// TIA Portal project "Text" (V21)

(* hardware
DEVICE "PLC_Text"  S7-1500 station
   slot 0: "Rail_0"  Rack  6ES7 590-1***0-0AA0
   slot 1: "PLC_Text"  CPU 1516-3 PN/DP  6ES7 516-3AN02-0AB0  V2.9
      slot 3: "CPU display_1"  6ES7591-1BA00-0AA0
      slot 32768: "PROFINET interface_1"  X1
         slot 32769: "Port_1"  X1 P1
         slot 32770: "Port_2"  X1 P2
      slot 33024: "PROFINET interface_2"  X2
         slot 33025: "Port_1"  X2 P1
      slot 33280: "DP interface_1"  X3
      slot 34817: "Virtual CP interface port_1"  Virtual CP interface port  Virtual CP interface port
*)

// ===== PLC "PLC_Text"  CPU 1516-3 PN/DP =====

VAR_GLOBAL   // PLC tag table "Beschriftung"
   "Lamp_Überlast" AT %Q0.0 : Bool;   // Überlast der Pumpe – Leuchte
   "Sensor_Niveau" AT %IW2 : Int;   // Capteur de niveau, en ‰
   "Etikett" AT %MW4 : Word;   // ラベル番号 (標識)
END_VAR

TYPE "typeLabel"
   STRUCT
      german : WString[40] := WSTRING#'Füllhöhe überschritten';   // Größe in Millilitern
      french : WString[40] := WSTRING#'Défaut de la vanne';   // Vanne fermée, ça bloque
      japanese : WString[20] := WSTRING#'液面センサー';   // 日本語のコメント
      chinese : WString[20] := WSTRING#'液位传感器';   // 中文注释
      plain : String[20] := 'It$'s 50% full';   // A quote and a percent sign
   END_STRUCT;
END_TYPE

DATA_BLOCK "Labels"   // DB1
TITLE = Beschriftungen für das Bedienfeld
{ S7_Optimized_Access := 'TRUE' }
VERSION : 0.1
   VAR
      current : "typeLabel";   // Die aktuelle Meldung
      list : Array[1..2] of "typeLabel";   // Zur Auswahl
      note : WString[40] := WSTRING#'Notiz: «Anführungszeichen»';   // Guillemets
   END_VAR
BEGIN
   list[1].german := WSTRING#'Ventil öffnet';
   list[2].japanese := WSTRING#'バルブが開く';
END_DATA_BLOCK

FUNCTION_BLOCK "Texts"   // FB1, SCL
TITLE = Überprüfung der Füllhöhe – ½ Liter
{ S7_Optimized_Access := 'TRUE' }
VERSION : 0.1
// Prüft die Füllhöhe. Vérifie le niveau. 液面を確認する。检查液位。
// A second comment line, with symbols: ± ° µ € ✓
   VAR_INPUT
      level : Real;   // Füllhöhe in ml – niveau de remplissage
      limit : Real := 500.0;   // Grenzwert ≥ 0
   END_VAR
   VAR_OUTPUT
      message : WString[60];   // Meldung für das Bedienfeld
      tooHigh : Bool;   // Zu hoch ✗
   END_VAR
   VAR
      label : "typeLabel";   // Texte in vier Sprachen
      path : String[40] := 'C:/data // not a comment';
      fake : String[40] := '(* not a comment either *)';
   END_VAR
BEGIN

    REGION Prüfung der Füllhöhe
        // Ist die Flasche zu voll? Est-elle trop pleine? 満杯ですか?
        #tooHigh := #level > #limit;
        IF #tooHigh THEN
            #message := #label.german;   // Deutsch zuerst
        ELSE
            #message := WSTRING#'Alles in Ordnung – OK';
        END_IF;
    END_REGION

    (* Ein Blockkommentar
       über zwei Zeilen: äöü ÄÖÜ ß *)
    #path := 'It$'s here: $'quoted$'';
END_FUNCTION_BLOCK